(* IEC 61131-3 sources: Caravan/Archiv/12-04-19/Stations/MachineControl/MachineControl/Class/_SIG_LSL_CMultimasterState, 1 file *)

(* ---- _SIG_LSL_CMultimasterState.st ---- *)
#include <.\LoaderItf.h>

(*!
<Class
	Name               = "_SIG_LSL_CMultimasterState"
	Revision           = "1.0"
	RealtimeTask       = "false"
	CyclicTask         = "false"
	BackgroundTask     = "false"
	Sigmatek           = "true"
	OSInterface        = "false"
	HighPriority       = "false"
	Automatic          = "false"
	UpdateMode         = "Prescan"
	SharedCommandTable = "true"
	Objectsize         = "(570,180)">
	<Channels>
		<Server Name="ClassSvr" Visualized="false" Initialize="false" WriteProtected="true" Retentive="false"/>
		<Server Name="PLC" Visualized="true" Initialize="false" WriteProtected="true" Retentive="false"/>
		<Server Name="Terminal" Visualized="true" Initialize="false" WriteProtected="true" Retentive="false"/>
	</Channels>
	<Dependencies>
		<Files>
			<File Path=".\LoaderItf.h" Include="true"/>
		</Files>
	</Dependencies>
</Class>
*)
_SIG_LSL_CMultimasterState : CLASS
	TYPE
	  _MMStateSvr :  //! <Type Public="true" Name="_MMStateSvr"/>
	  (
	    Offline:=0,  //! <Type Comment="Station offline." Name="_MMStateSvr.Offline"/>
	    Online_Initializing:=1,  //! <Type Comment="Station online,&#10;servers not updated." Name="_MMStateSvr.Online_Initializing"/>
	    Online:=2,  //! <Type Comment="Station online,&#10;all servers existing and initalized." Name="_MMStateSvr.Online"/>
	    Online_NotAllServerAvailable:=3,  //! <Type Comment="Station online,&#10;not all server exists, existing servers initalized." Name="_MMStateSvr.Online_NotAllServerAvailable"/>
	    SvrNotFoundAtStation:=16  //! <Type Comment="No valid LasalID for server found." Name="_MMStateSvr.SvrNotFoundAtStation"/>
	  )$UDINT;
	END_TYPE
  //Servers:
	ClassSvr 	: SvrChCmd_DINT;
	Terminal 	: SvrCh__MMStateSvr_PTofCls__SIG_LSL_CMultimasterState;
	PLC 	: SvrCh__MMStateSvr_PTofCls__SIG_LSL_CMultimasterState;
  //Clients:
  //Variables:
		m_arrSERVERS : ARRAY [0..255] OF ^_MMStateSvr;

  //Functions:

	FUNCTION _SIG_LSL_CMultimasterState
		VAR_OUTPUT
			ret_code 	: ConfStates;
		END_VAR;

	FUNCTION GLOBAL Callback
		VAR_INPUT
			pThis 	: ^void;
			udStationId 	: UDINT;
			szStationName 	: ^CHAR;
			udServerHandle 	: UDINT;
			szServerName 	: ^CHAR;
			udState 	: _SIG_LSL_CMultimasterState::_MMStateSvr;
		END_VAR;

	FUNCTION VIRTUAL GLOBAL UserCallback
		VAR_INPUT
			udStationId 	: UDINT;
			szStationName 	: ^CHAR;
			udServerHandle 	: UDINT;
			szServerName 	: ^CHAR;
			udState 	: _SIG_LSL_CMultimasterState::_MMStateSvr;
		END_VAR;
  //Tables:
	FUNCTION @STD
		VAR_OUTPUT
			ret_code	: CONFSTATES;
		END_VAR;
	FUNCTION GLOBAL TAB @CT_;
END_CLASS;

FUNCTION GLOBAL _SIG_LSL_CMultimasterState::Callback
VAR_INPUT
  pThis           : ^void;
  udStationId     : UDINT;
  szStationName   : ^CHAR;
  udServerHandle	 : UDINT;
  szServerName  	: ^CHAR;
  udState 	      : _SIG_LSL_CMultimasterState::_MMStateSvr;
END_VAR
  this := pThis$^_SIG_LSL_CMultimasterState;

  if ( udState$UDINT < __MMSTATE_SERVER_BEGIN_ ) then
    if ( m_arrSERVERS[TO_USINT(udStationId)] <> NIL ) then
      m_arrSERVERS[TO_USINT(udStationId)]^ := ( udState );
    end_if;

  end_if;

  UserCallback(udStationId, szStationName, udServerHandle, szServerName, udState);
END_FUNCTION

#pragma warning(disable:73);
FUNCTION VIRTUAL GLOBAL _SIG_LSL_CMultimasterState::UserCallback
VAR_INPUT
  udStationId     : UDINT;
  szStationName   : ^CHAR;
  udServerHandle	 : UDINT;
  szServerName  	: ^CHAR;
  udState 	      : _SIG_LSL_CMultimasterState::_MMStateSvr;
END_VAR
END_FUNCTION
#pragma warning(default:73);

FUNCTION _SIG_LSL_CMultimasterState::_SIG_LSL_CMultimasterState
VAR_OUTPUT
  ret_code 	: ConfStates;
END_VAR
    ret_code := C_OK;

    //for each MM-Station a entry in ARRAY for faster access:
    _memset(#m_arrSERVERS[0], 0, SIZEOF(m_arrSERVERS));
    m_arrSERVERS[TO_USINT(LDR_MM_StatNameGetNr("Terminal"))] := #Terminal$_MMStateSvr;
    m_arrSERVERS[TO_USINT(LDR_MM_StatNameGetNr("PLC"))] := #PLC$_MMStateSvr;
    //Install callback at Loader:
    LDR_MM_InstallCallback(#Callback(), this);

END_FUNCTION
